// TIA Portal V21 export
// export: Created 2026-11-10T19:16:32.7469358Z, ExportSetting WithDefaults, DisplayName Totally Integrated Automation Portal, DisplayVersion V21 Update 3, DisplayName STEP 7 Professional, DisplayVersion V21 Update 3, DisplayName STEP 7 Safety, DisplayVersion V21, DisplayName Tech WebApplication, DisplayVersion V21, DisplayName WinCC Basic/Comfort/Advanced, DisplayVersion V21 Update 3, DisplayName WinCC Unified, DisplayVersion V21 Update 3
DATA_BLOCK "DB_300"   // DB1
VERSION : 0.1
// stored: AutoNumber true, IsOnlyStoredInLoadMemory false, IsWriteProtectedInAS false
   VAR RETAIN
      x : Bool;
      i : Int := 30;
      d : DInt;
      r : Real := 1.25;
      t : Time;
      dtv : Date_And_Time;
      s : String[8] := 'S7-300';
      arr : Array[0..3] of Int;
      "m" : Array[0..1, 0..1] of Word;
      st : Struct
         p : Word;
         q : Byte;
      END_STRUCT;
      u { S7_SetPoint := 'True'} : "UDT_300";
   END_VAR
BEGIN
   arr[2] := 22;
   "m"[1,1] := WORD#16#ABCD;
END_DATA_BLOCK
